INTERFACE ITF_Banddepalletizer

METHOD Aborted : BOOL
VAR_INPUT
END_VAR
END_METHOD

METHOD Aborting : BOOL
VAR_INPUT
END_VAR
END_METHOD

METHOD Clearing : BOOL
VAR_INPUT
END_VAR
END_METHOD

METHOD Execute : BOOL
VAR_INPUT
END_VAR
END_METHOD

METHOD Held : BOOL
VAR_INPUT
END_VAR
END_METHOD

METHOD Holding : BOOL
VAR_INPUT
END_VAR
END_METHOD

METHOD Idle : BOOL
VAR_INPUT
END_VAR
END_METHOD

METHOD Resetting : BOOL
VAR_INPUT
END_VAR
END_METHOD

METHOD Starting : BOOL
VAR_INPUT
END_VAR
END_METHOD

METHOD Stopped : BOOL
VAR_INPUT
END_VAR
END_METHOD

METHOD Stopping : BOOL
VAR_INPUT
END_VAR
END_METHOD

METHOD Suspended : BOOL
VAR_INPUT
END_VAR
END_METHOD

METHOD Suspending : BOOL
VAR_INPUT
END_VAR
END_METHOD

METHOD Unholding : BOOL
VAR_INPUT
END_VAR
END_METHOD

METHOD Unsuspending : BOOL
VAR_INPUT
END_VAR
END_METHOD

END_INTERFACE

(* stored: Version 1.1.0.1
   Itf ITF_Banddepalletizer: Id {b09bf2ba-d668-46e6-a510-ea61c886fdd7}
   Folder Methods: Id {e7934a6e-4fbf-45cc-9392-559bfdf7288e}
   Method Aborted: Id {d259aaac-ef8e-4ef9-9913-9e4718b0fb37}
   Method Aborting: Id {ff4e62dc-5e0c-4abe-87b1-df5734a3d4b7}
   Method Clearing: Id {c1bf0531-9200-43fb-8180-3f0554778ea2}
   Method Execute: Id {613ce1b5-979e-42fb-9ab7-1900e07fc1b8}
   Method Held: Id {a6b506ab-6802-4462-be53-7c8f91be1104}
   Method Holding: Id {5b585d67-fc1c-4124-a13a-8908ca228e17}
   Method Idle: Id {474d33b2-bac7-4686-8319-c49324562eba}
   Method Resetting: Id {fb4373f8-f768-4d13-ad43-7de8c374b656}
   Method Starting: Id {7cb9b9b6-b2d5-445b-a646-1ae8e325ab0f}
   Method Stopped: Id {8dba2f31-d754-4556-aa2d-7be68ee1b7f7}
   Method Stopping: Id {569a5c14-f918-4955-8090-eb2fb6b4b935}
   Method Suspended: Id {1a41f243-83c2-4f81-ba73-117cc67690c6}
   Method Suspending: Id {8db35fa5-54bc-4b08-86c0-69939833a91e}
   Method Unholding: Id {404c7e3f-47aa-47dc-a08d-40dac1fbade1}
   Method Unsuspending: Id {b846eb73-8b1b-49da-a0f7-6f9baab539ef} *)
